FUNCTION_BLOCK FB_LineClamp IMPLEMENTS I_LineClamp
VAR_INPUT
    Jammed : BOOL;
END_VAR
VAR
    Position : DINT;
END_VAR

METHOD Follow : DINT
VAR_INPUT
    Extend : BOOL;
END_VAR
IF NOT Extend THEN Position := MAX(0, Position - 4);
ELSIF NOT Jammed THEN Position := MIN(16, Position + 4);
END_IF
Follow := Position;
END_METHOD

METHOD Home
Position := 0;
END_METHOD

END_FUNCTION_BLOCK

(* stored: Version 1.1.0.1
   POU FB_LineClamp: Id {CB31703C-BDF0-4A15-AF15-000000000006}
   Method Follow: Id {CB31703C-BDF0-4A15-AF15-000000000004}
   Method Home: Id {CB31703C-BDF0-4A15-AF15-000000000005} *)
